// TIA Portal V20 export
// export: Created 2026-10-19T18:07:16.0439433Z, ExportSetting WithDefaults, DisplayName Totally Integrated Automation Portal, DisplayVersion V20 Update 6, DisplayName TIA Portal Openness, DisplayVersion V20 Update 6, DisplayName TIA Portal Version Control Interface, DisplayVersion V20 Update 6, DisplayName SINAMICS Startdrive Advanced, DisplayVersion V20 SP1, DisplayName SINAMICS Startdrive G130, G150, S120, S150, SINAMICS MV, G220, S200, S210, DisplayVersion V20 SP1, DisplayName SINAMICS Startdrive G110M, G120, G120C, G120D, G120P, G115D, DisplayVersion V20 SP1, DisplayName STEP 7 Professional, DisplayVersion V20 Update 6, DisplayName STEP 7 Safety, DisplayVersion V20 Update 2, DisplayName WinCC Basic/Comfort/Advanced, DisplayVersion V20 Update 6, DisplayName WinCC Unified, DisplayVersion V20 Update 6
DATA_BLOCK "Watchdog_Settings"   // DB134
{ S7_Optimized_Access := 'TRUE' }
VERSION : 0.1
// stored: AutoNumber true, DBAccessibleFromOPCUA true, DBAccessibleFromWebserver true, InstanceOfName Watchdog_Settings_UDT, InstanceOfType UDT, IsOnlyStoredInLoadMemory false, IsWriteProtectedInAS false
"Watchdog_Settings_UDT"
   // VAR
   //    Cnv_Entry : UDInt := 500;
   //    Cnv_PopUp : Array[1..4] of UDInt;
   //    Cnv_Exit : UDInt := 500;
   //    VTD : UDInt := 500;
   //    EConveyor : UDInt := 500;
   //    Cnv_Buffer : Array[1..3] of UDInt;
   //    Roller_TO_Roller : UDInt := 500;
   //    Chain_TO_Chain : UDInt := 500;
   //    Pop4_TO_Pick : UDInt := 500;
   //    Pick_TO_Pop1 : UDInt := 500;
   //    Weigh_Station : UDInt := 500;
   //    Profile_Station : UDInt := 500;
   //    Pallet_INOut : UDInt := 500;
   //    Shuttle_INOut : UDInt := 500;
   // END_VAR
BEGIN
   Cnv_PopUp[1..4] := 500;
   Cnv_Buffer[1..3] := 500;
END_DATA_BLOCK
